(* PLC project fbd_fan_damper_bomb, Anonymous Benchmark Suite 1.0 *)
(* stored: creationDateTime 2026-08-26T00:00:00 *)

PROGRAM air_handler
  VAR_INPUT
    fan_cmd : BOOL;
    damper_open : BOOL;
    smoke : BOOL;
  END_VAR
  VAR_OUTPUT
    fan : BOOL;
  END_VAR

(* FBD diagram, written out as Structured Text *)
fan := fan_cmd AND NOT smoke;
END_PROGRAM

CONFIGURATION Config0
  RESOURCE Res0 ON PLC
    TASK tcyclic(INTERVAL := T#10ms, PRIORITY := 0);
    PROGRAM inst0 WITH tcyclic : air_handler;
  END_RESOURCE
END_CONFIGURATION
